FUNCTION_BLOCK T_TestDirectory
VAR
  createDirectory : FB_CreateDir;
  requested : BOOL;
  _ready : BOOL;
END_VAR

IF _ready THEN
  RETURN;
END_IF

createDirectory(sNetId := '', sPathName := TestFiles.DIRECTORY, bExecute := TRUE);

IF requested AND NOT createDirectory.bBusy THEN
  _ready := TRUE;
END_IF

requested := TRUE;

PROPERTY Ready : BOOL
GET
Ready := _ready;
END_GET
END_PROPERTY

END_FUNCTION_BLOCK

(* stored: Version 1.1.0.1, ProductVersion 3.1.4026.25
   POU T_TestDirectory: Id {3a67114a-7265-4ca9-9903-10d074580a63}, SpecialFunc None
   Property Ready: Id {7f37cdd5-a72d-4c53-998e-557cde053969}
   Get Get: Id {e3c9d33e-9001-4f03-a18e-1ff14ecbc40f} *)
